# EPICS substitutions: db/Beckhoff_7XXX/ecmcEX72XX_OPT_info2Errors.substitutions
file "ecmcEX72XX_OPT_errors.template"
{
  pattern {CH_ID}
          {"$(OPT_CH_ID=01)"}
}
